// TIA Portal V19 export
TYPE "PID"
   STRUCT
      P : Real;
      I : Real;
      D : Real;
   END_STRUCT;
END_TYPE
